(*
SPDX-FileCopyrightText: © 2026 Oleksandr Tiutyk <trofimich@gmail.com>
SPDX-License-Identifier: MIT
License: https://opensource.org/license/mit
*)

(*!
<summary>Provides DATE_AND_TIME limits and date/time formatting with selectable separators.</summary>
<description>
Formatting removes the type prefix from the native text representation. Each separator can contain one
character or be empty to omit that separator. No time-zone conversion is performed.
</description>
*)

{attribute 'no_explicit_call' := 'Direct call is not allowed'}
PROGRAM DateAndTimes
VAR CONSTANT
	MIN_VALUE : DATE_AND_TIME := DT#1970-1-1-0:0:0;
	MAX_VALUE : DATE_AND_TIME := DT#2106-02-07-06:28:15;
END_VAR
VAR
	{attribute 'hide'} 
	_ClassName : STRING := __POUNAME();
END_VAR

{attribute 'monitoring' := 'call'}
PROPERTY ClassName : REFERENCE TO STRING
GET
ClassName REF= _ClassName;
END_GET
END_PROPERTY

(*!
<summary>Provides the library namespace used in diagnostics.</summary>
<description>
Borrowed read-only reference to the compiler-initialized library namespace; no ownership transfer.
</description>
*)
{attribute 'monitoring' := 'call'}
PROPERTY NamespaceName : REFERENCE TO STRING
GET
NamespaceName REF= CurrentNamespace.Name;
END_GET
END_PROPERTY

(*!
<summary>Formats the date and time without the type prefix, using the supplied separators.</summary>
<description>
Empty separators remove the corresponding delimiters. Date and time fields retain their native order and
padding; any fractional-second suffix is preserved.
</description>
*)
//!<param name="value">Date and time to format without time-zone conversion.</param>
//!<param name="dateValuesSeparator">Separator between year, month and day; empty omits both delimiters.</param>
//!<param name="dateAndTimeSeparator">Separator between date and time; empty omits it.</param>
//!<param name="timeValuesSeparator">Separator between hours, minutes and seconds; empty omits both delimiters.</param>
METHOD ToString : STRING
VAR_INPUT
	value : DATE_AND_TIME;
	dateValuesSeparator : STRING(1) := '_';
	dateAndTimeSeparator : STRING(1) := '-';
	timeValuesSeparator : STRING(1) := '_';
END_VAR
ToString := TO_STRING(value);

ToString := Tc2_Standard.DELETE(STR := ToString, LEN := 3, POS := 1);

(* Replace from right to left so empty separators do not shift pending positions. *)
ToString := Tc2_Standard.REPLACE(STR1 := ToString, STR2 := timeValuesSeparator, L := 1, P := 17);
ToString := Tc2_Standard.REPLACE(STR1 := ToString, STR2 := timeValuesSeparator, L := 1, P := 14);
ToString := Tc2_Standard.REPLACE(STR1 := ToString, STR2 := dateAndTimeSeparator, L := 1, P := 11);
ToString := Tc2_Standard.REPLACE(STR1 := ToString, STR2 := dateValuesSeparator, L := 1, P := 8);
ToString := Tc2_Standard.REPLACE(STR1 := ToString, STR2 := dateValuesSeparator, L := 1, P := 5);
END_METHOD

(*!
<summary>Formats the date and time without the type prefix, using the supplied separators.</summary>
<description>
Empty separators remove the corresponding delimiters. Date and time fields retain their native order and
padding; any fractional-second suffix is preserved.
</description>
*)
//!<param name="value">Date and time to format without time-zone conversion.</param>
//!<param name="dateValuesSeparator">Separator between year, month and day; empty omits both delimiters.</param>
//!<param name="dateAndTimeSeparator">Separator between date and time; empty omits it.</param>
//!<param name="timeValuesSeparator">Separator between hours, minutes and seconds; empty omits both delimiters.</param>
METHOD ToWideString : WSTRING
VAR_INPUT
	value : DATE_AND_TIME;
	dateValuesSeparator : WSTRING(1) := "_";
	dateAndTimeSeparator : WSTRING(1) := "-";
	timeValuesSeparator : WSTRING(1) := "_";
END_VAR
ToWideString := TO_WSTRING(value);

ToWideString := Tc2_Standard.WDELETE(STR := ToWideString, LEN := 3, POS := 1);

(* Replace from right to left so empty separators do not shift pending positions. *)
ToWideString := Tc2_Standard.WREPLACE(STR1 := ToWideString, STR2 := timeValuesSeparator, L := 1, P := 17);
ToWideString := Tc2_Standard.WREPLACE(STR1 := ToWideString, STR2 := timeValuesSeparator, L := 1, P := 14);
ToWideString := Tc2_Standard.WREPLACE(STR1 := ToWideString, STR2 := dateAndTimeSeparator, L := 1, P := 11);
ToWideString := Tc2_Standard.WREPLACE(STR1 := ToWideString, STR2 := dateValuesSeparator, L := 1, P := 8);
ToWideString := Tc2_Standard.WREPLACE(STR1 := ToWideString, STR2 := dateValuesSeparator, L := 1, P := 5);
END_METHOD

END_PROGRAM

(* stored: Version 1.1.0.1
   POU DateAndTimes: Id {0483a592-4912-4994-8cc7-7285a0ab6a20}, SpecialFunc None
   Property ClassName: Id {6f3d40ea-0adf-43e0-9f6c-bb2b4322828f}
   Get Get: Id {79a6c653-6fbb-470a-9071-7d181520f68d}
   Property NamespaceName: Id {dc154108-24f4-48b1-8479-bc7faf5bd8ee}
   Get Get: Id {fa3a7606-7124-42f1-be10-98cd079db160}
   Method ToString: Id {e0790e93-eb77-4ac6-a5e7-38f9fddb40f4}
   Method ToWideString: Id {7498afc1-9ae1-4986-8ff2-63e14a92dea2} *)
